Fanuc KAREL source: KT00197.KL

PROGRAM KT00197
%NOLOCKGROUP
VAR
  B1: BOOLEAN
  Y2: ARRAY[2] OF BYTE
  OUT: BOOLEAN
BEGIN
  B1 = TRUE
    Y2[1] = 3
  OUT = B1 AND Y2[1]
END KT00197
